// TIA Portal V19 export
// export: Created 2026-10-15T09:44:22.9560565Z, ExportSetting WithDefaults, DisplayName Totally Integrated Automation Portal, DisplayVersion V19, DisplayName TIA Portal Openness, DisplayVersion V19, DisplayName TIA Portal Version Control Interface, DisplayVersion V19, DisplayName STEP 7 Professional, DisplayVersion V19, DisplayName STEP 7 Safety, DisplayVersion V19, DisplayName WinCC Basic/Comfort/Advanced, DisplayVersion V19, DisplayName WinCC Unified, DisplayVersion V19
FUNCTION "ROLL_GetDW" : Word   // FC3, SCL
{ S7_Optimized_Access := 'TRUE' }
VERSION : 0.1
// stored: AutoNumber true, IsIECCheckEnabled false, SetENOAutomatically false, UDAEnableTagReadback false
   VAR_INPUT
      DbNumber : Int;
      Index : Int;
   END_VAR
BEGIN

   #ROLL_GetDW := W#16#0000;
   IF (#Index < 0) OR (#Index > 131) THEN
       "ROLL_IO".ConversionFault := TRUE;
       RETURN;
   END_IF;
   CASE #DbNumber OF
       15:
           #ROLL_GetDW := "ROLL_DB15".DW[#Index];
       19:
           #ROLL_GetDW := "ROLL_DB19".DW[#Index];
       ELSE
           "ROLL_IO".ConversionFault := TRUE;
   END_CASE;
END_FUNCTION
